(* IEC 61131-3 sources: codesys-api/examples/plc_architecture/bench/st_native, 2 files *)

(* ---- PRG_NativeSerial.st ---- *)
PROGRAM PRG_NativeSerial
// Bench, --serial native (generated from bench/st_native): the PLC's RJ12 port is polled by the device tree's
// Modbus_COM master, one server per unit, each channel mapped to GVL_Native.Unit<n>. Called in the bus task
// (the bus cycle task, which refreshes those images): hands each image to the same decode table as the
// ModbusFB lines and turns the server's xError into source health. The device tree gives no per-reply event,
// so SourceLastGoodMs means "no error flagged as of this cycle", not "a reply arrived". And xError only
// describes the latest poll: with auto-restart a dead server's flag clears at every retry (bench, 2026-10-20:
// unit 5 silent, healthy in a third of control scans with its last image), so a server counts as healthy only
// after HOLD_MS without an error.
VAR CONSTANT
	HOLD_MS : ULINT := 2500;            // longer than a channel cycle plus the reply timeout
END_VAR
VAR
	Words : ARRAY[0..124] OF WORD;
	Bits : ARRAY[0..1999] OF BYTE;
	WasError : ARRAY[1..@@COUNT@@] OF BOOL;
	ErrorEdges : ARRAY[1..@@COUNT@@] OF UDINT;     // diagnostics: times each server went into error
	ErrorCycles : ARRAY[1..@@COUNT@@] OF UDINT;    // ... and bus cycles it spent in error (share = / CycleCount)
	CycleCount : UDINT;
	LastErrorMs : ARRAY[1..@@COUNT@@] OF ULINT;
	NowMs : ULINT;
END_VAR
// ---- implementation ----
NowMs := F_NowMs();
CycleCount := CycleCount + 1;
@@CALLS@@

(* ---- PRG_NativeSerial.Take.st ---- *)
METHOD Take : BOOL
// One server: decode its image into GVL_Bus.Raw once it has been error-free for HOLD_MS; unhealthy until then.
VAR_INPUT
	Number : INT;                       // position in WasError / ErrorEdges
	Block : INT;                        // its GVL_Bus.Blocks row (the decode description)
	IsError : BOOL;                     // the server's xError
END_VAR
VAR_IN_OUT
	Image : ARRAY[0..5] OF WORD;
END_VAR
VAR
	Source : INT;
	Index : INT;
END_VAR
// ---- implementation ----
Source := GVL_Bus.Blocks[Block].Source;
IF IsError AND NOT WasError[Number] THEN
	ErrorEdges[Number] := ErrorEdges[Number] + 1;
END_IF
WasError[Number] := IsError;
IF IsError THEN
	ErrorCycles[Number] := ErrorCycles[Number] + 1;
	LastErrorMs[Number] := NowMs;
END_IF
GVL_Bus.SourceWriting[Source] := TRUE;
IF LastErrorMs[Number] <> 0 AND NowMs - LastErrorMs[Number] < HOLD_MS THEN
	GVL_Bus.SourceHealthy[Source] := FALSE;
ELSE
	FOR Index := 0 TO 5 DO
		Words[Index] := Image[Index];
	END_FOR
	F_BusDecode(FirstEntry := GVL_Bus.Blocks[Block].FirstEntry, EntryCount := GVL_Bus.Blocks[Block].EntryCount,
		Words := Words, Bits := Bits);
	GVL_Bus.SourceHealthy[Source] := TRUE;
	GVL_Bus.SourceLastGoodMs[Source] := NowMs;
END_IF
GVL_Bus.SourceWriting[Source] := FALSE;
Take := TRUE;
